Fanuc KAREL source: kt00344.KL

-- PROVISIONAL review KL for V770-1; original PC SHA256 e815b5f9bbd82aa66e93eaaa5c79ccb7f75c281742c777fbd439a348b916e198
-- Incomplete behavior may be omitted. Consult companion uncertainty JSON. Do not deploy.
PROGRAM KT00344
%NOLOCKGROUP
VAR
  R2 : REAL
  OUT : BOOLEAN
-- UNRESOLVED_DECL H1 type=002017
BEGIN
  -- UNRESOLVED_PC offsets 5-19; opcodes 2E,22,9D,33,B4
  -- UNRESOLVED_PC offsets 24-35; opcodes 2E,23
  -- UNRESOLVED_PC offsets 40-65; opcodes 22,9D,33,B3,21,29,64,29,6F,23
  -- UNRESOLVED_PC offsets 70-74; opcodes 7F
END KT00344
